// TIA Portal V20 export
// export: Created 2026-10-12T04:58:21.888491Z, ExportSetting WithDefaults, DisplayName Totally Integrated Automation Portal, DisplayVersion V20, DisplayName TIA Portal Openness, DisplayVersion V20, DisplayName TIA Portal Teamcenter Gateway, DisplayVersion V20, DisplayName TIA Portal Version Control Interface, DisplayVersion V20, DisplayName SINAMICS Startdrive Advanced, DisplayVersion V20 SP1 Update 2, DisplayName SINAMICS Startdrive G110M, G120, G120C, G120D, G120P, G115D, DisplayVersion V20 SP1 Update 2, DisplayName SINAMICS Startdrive G130, G150, S120, S150, SINAMICS MV, G220, S200, S210, DisplayVersion V20 SP1 Update 2, DisplayName STEP 7 Professional, DisplayVersion V20, DisplayName STEP 7 Safety, DisplayVersion V20, DisplayName WinCC Basic/Comfort/Advanced, DisplayVersion V20, DisplayName WinCC Professional, DisplayVersion V20, DisplayName WinCC Unified, DisplayVersion V20
FUNCTION "FRK_SetValidateEnd" : Bool   // FC115, SCL
{ S7_Optimized_Access := 'TRUE' }
VERSION : 0.1
// stored: AutoNumber true, IsIECCheckEnabled false, SetENOAutomatically false, UDAEnableTagReadback false
   VAR_INPUT
      RootIndex : Int;
   END_VAR
   VAR_TEMP
      Index : Int;
   END_VAR
BEGIN

   #FRK_SetValidateEnd := FALSE;
   FOR #Index := 1 TO "FRK_SetRuntime".Work[#RootIndex].Payload.Info.RecordCount DO
       IF NOT "FRK_SetRuntime".Work[#RootIndex].Seen[#Index] THEN
           "FRK_SetRuntime".Work[#RootIndex].RejectScope := "FRK_SetRuntime".Work[#RootIndex].Payload.Records[#Index].Scope;
           "FRK_SetRuntime".Work[#RootIndex].RejectKey := "FRK_SetRuntime".Work[#RootIndex].Payload.Records[#Index].WriteKey;
           RETURN;
       END_IF;
   END_FOR;
   #FRK_SetValidateEnd := "FRK_SetRuntime".Work[#RootIndex].Matched = "FRK_SetRuntime".Work[#RootIndex].Payload.Info.RecordCount;
END_FUNCTION
